ABB RAPID module: TgtProg.mod

MODULE MainModule
GLOBAL VAR robtarget robpoint0= p:{{-607.850, 543.849, 363.215},{0.374108, 0.285846, 0.853660, -0.222712}}{cfg 0,0,0,0}{7.000000,0.0,0.0,0.0,0.0,0.0}

GLOBAL Proc main()
    MoveL robpoint0,v50,z50,tool03,wobj16
EndProc
EndModule
